// TIA Portal V21 export
// export: Created 2026-11-10T19:16:29.3875875Z, ExportSetting WithDefaults, DisplayName Totally Integrated Automation Portal, DisplayVersion V21 Update 3, DisplayName STEP 7 Professional, DisplayVersion V21 Update 3, DisplayName STEP 7 Safety, DisplayVersion V21, DisplayName Tech WebApplication, DisplayVersion V21, DisplayName WinCC Basic/Comfort/Advanced, DisplayVersion V21 Update 3, DisplayName WinCC Unified, DisplayVersion V21 Update 3
DATA_BLOCK "DB_12Opt"   // DB1
{ S7_Optimized_Access := 'TRUE' }
VERSION : 0.1
// stored: AutoNumber true, DBAccessibleFromOPCUA true, IsOnlyStoredInLoadMemory false, IsRetainMemResEnabled false, IsWriteProtectedInAS false, MemoryReserve 100
   VAR
      x : Bool;
      i : Int := 12;
      d : DInt;
      r : Real;
      lr : LReal;
      t : Time;
      dtl : DTL;
      s : String[10] := 'S7-1200';
      ws : WString;
      a2 : Array[0..1, 0..2] of Int;
      st : Struct
         p : Word;
         q : Array[1..3] of Byte;
      END_STRUCT;
      u { S7_SetPoint := 'True'} : "UDT_12";
      au { S7_SetPoint := 'True'} : Array[0..1] of "UDT_12";
      tm { S7_SetPoint := 'True'} : IEC_TIMER;
   END_VAR
   VAR RETAIN
      rr : UDInt;
   END_VAR
BEGIN
   a2[1,2] := 7;
   u."b" := 2.5;
   au[1]."a" := 9;
END_DATA_BLOCK
